ORGANIZATION_BLOCK "Main"
{ S7_Optimized_Access := 'TRUE' }
VERSION : 0.1
BEGIN
    "GDB_OperationsTest"();
    "FRK_TestPublish"(Complete := "GDB_OperationsTest".Done, Image0 := DWORD#3497805631, Image1 := DWORD#611401252, Image2 := DWORD#132661567, Image3 := DWORD#130345828, Image4 := DWORD#4112764091, Image5 := DWORD#1815743570, Image6 := DWORD#575805802, Image7 := DWORD#101359597, Result := "GDB_OperationsTest".Result, Status := "GDB_OperationsResultTest".Status);
END_ORGANIZATION_BLOCK
